Fanuc KAREL source: kb00087.KL

PROGRAM KB00087
%NOLOCKGROUP
%ENVIRONMENT REGOPE
VAR
P1:INTEGER;P2:INTEGER;RESULT : XYZWPREXT
BEGIN
--
--
P1=1
P2=1
RESULT=GET_POS_REG(P1,P2,1)
END KB00087
